TYPE ET_SpindleCtrl :
(
	ET_SpindleCtrl_eWaitExecute := 0,
	ET_SpindleCtrl_eCtrlEnable := 5,
	ET_SpindleCtrl_eWfCtrlEnabled := 10,
	ET_SpindleCtrl_eSpindleStop := 15,
	ET_SpindleCtrl_eWfSpindleStopped := 20,
	ET_SpindleCtrl_eSpindleRun := 25,
	ET_SpindleCtrl_eWfSpindleRunning := 30,
	ET_SpindleCtrl_eDone := 197,
	ET_SpindleCtrl_eError := 198,
	ET_SpindleCtrl_eNoExecute := 199
);
END_TYPE

(* stored: Version 1.1.0.1, ProductVersion 3.1.4024.15
   DUT ET_SpindleCtrl: Id {f0db0bd1-4976-4345-89ba-c3b8649cf54d} *)
